(* IEC 61131-3 sources: 2026_Projet_YGO_ExcavatriceDragage/CODE/H_TREUILS_BENNE, 13 files *)

(* ---- FB_BucketCmdArbitration.st ---- *)
(* ═══════════════════════════════════════════════════════════════
   🪣 FB_BucketCmdArbitration — Arbitrage de commande benne
   ───────────────────────────────────────────────────────────────
   🎯 Rôle : Arbitrer la source de commande benne (boutons IHM /
       séquencement couplé both / demande cycle selon le mode) et produire
       les commandes arbitrées (ouverture, fermeture, contacteur Kobold).
   🔌 FB d'arbitrage (non-mouvement) : ne porte ni SafeStop ni StartStop
       de sécurité — il produit la commande logique, la safety reste dans
       FB_Bucket / FB_Safety_Winch.
   📄 Doc : DOC/AF/AF_Partie-10_Fonction_Winch_v2.1.md
   🔒 Bit-identique à l'ancien PRG_04 §1/§2 (refactor POO §5 : décision dans
       le FB, plus dans le PRG). Symétrique à FB_WinchCmdArbitrationM1/M2.
   ═══════════════════════════════════════════════════════════════ *)

FUNCTION_BLOCK FB_BucketCmdArbitration
VAR_INPUT
    Enable    : BOOL;  // --> [CMD] Autorisation FB (TRUE=arbitre actif)
    Auth      : ST_Modes_Autorisations;          // --> [CMD] Autorisations mode (Mode, gating séquencement couplé)
    ReqBucket : ST_ProgramBucketRequest;            // --> [REQ] Demande cycle benne (SEMI_AUTO)
    IHM       : ST_fbBucketCmdArbitration_IHM;      // --> [CMD] Boutons IHM benne (BtnOpen/BtnClose)
    Context   : ST_fbBucketCmdArbitration_Context;   // --> [STAT] Gating séquencement couplé benne
END_VAR
VAR_OUTPUT
    Ready     : BOOL;  // <-- [STAT] FB prêt à arbitrer (Enable)
    CmdOpen_IHM  : BOOL;  // <-- [CMD] Commande ouverture benne arbitrée
    CmdClose_IHM : BOOL;  // <-- [CMD] Commande fermeture benne arbitrée
    KoboldContactorCmdArbitrated : BOOL;  // <-- [CMD] Ordre contacteur capteur fond Kobold arbitré
    WinchBothDiveBucketOpenArmed    : BOOL;  // <-- [STAT] Séquencement couplé : descente benne ouverte armé
    WinchBothAscentBucketCloseArmed : BOOL;  // <-- [STAT] Séquencement couplé : montée benne fermée armé
END_VAR

// === IMPLEMENTATION ===

Ready := Enable;

IF NOT Enable THEN
    CmdOpen_IHM  := FALSE;
    CmdClose_IHM := FALSE;
    KoboldContactorCmdArbitrated := FALSE;
    WinchBothDiveBucketOpenArmed    := FALSE;
    WinchBothAscentBucketCloseArmed := FALSE;
ELSE
    // ── Règle absolue en pilotage both normal (bit-identique PRG_04 §1) ──
    // Descente autorisée UNIQUEMENT benne ouverte, montée UNIQUEMENT benne fermée.
    // T248 : une fois la phase couplée VERROUILLÉE (benne amenée dans l'état requis pour
    // ce maintien joystick), on n'arme plus dive-open / ascent-close -> la perte de
    // l'état ouvert/fermé EN MOUVEMENT ne relance aucune correction benne et ne bloque
    // plus le mouvement couplé ("descente/montée interdite" fantôme).
    WinchBothDiveBucketOpenArmed := Context.TglEnableCoupledBucketSequencing
        AND (Auth.Mode <> E_Mode.SEMI_AUTO)
        AND NOT Context.CoupledPhaseLocked
        AND Context.MotionActive AND Context.ReqDescend
        AND NOT Context.BucketIsOpen;
    WinchBothAscentBucketCloseArmed := Context.TglEnableCoupledBucketSequencing
        AND (Auth.Mode <> E_Mode.SEMI_AUTO)
        AND NOT Context.CoupledPhaseLocked
        AND Context.MotionActive AND Context.ReqAscent
        AND NOT Context.BucketIsClosed;

    // ── Ouverture benne : bouton IHM OU séquencement couplé descente benne ouverte
    //    OU demande cycle (bit-identique PRG_04 §2) ──
    CmdOpen_IHM := IHM.BtnOpen OR WinchBothDiveBucketOpenArmed OR ReqBucket.ReqOpen;

    // ── Fermeture benne : demande cycle > séquencement couplé montée benne fermée
    //    > bouton IHM (bit-identique PRG_04 §1) ──
    IF ReqBucket.ReqClose THEN
        CmdClose_IHM := TRUE;
    ELSIF WinchBothAscentBucketCloseArmed THEN
        CmdClose_IHM := TRUE;
    ELSE
        CmdClose_IHM := IHM.BtnClose;
    END_IF;

    // ── Contacteur Kobold : demande cycle (source unique PRG_03, bit-identique PRG_04 §1) ──
    KoboldContactorCmdArbitrated := ReqBucket.ReqKoboldMeasureEnable;
END_IF;

END_FUNCTION_BLOCK

(* ---- FB_DriftGuard.st ---- *)
(* =======================================================================
   📐 FB_DriftGuard — Détection de dérive de position sous armement
   ───────────────────────────────────────────────────────────────
   🎯 Rôle : Capture position de référence et détection de dérive anormale
   📄 Doc métier : DOC/AF/AF_Partie-10_Fonction_Winch_v2.1.md
   🔌 Interface : Brique interne de sécurité (compose FB_Safety_Winch)
   🔒 Sécurité : Détection de mouvement non commandé et glissement
   ======================================================================= *)

FUNCTION_BLOCK PUBLIC FB_DriftGuard
VAR_INPUT
    // === COMMANDES ET SEUILS ===
    Arm                             : BOOL;                           // --> [CMD] Condition d'armement de la surveillance
    PositionM                       : REAL;                           // --> [HW] Position courante a surveiller (m)
    ToleranceM                      : REAL;                           // --> [CFG] Tolerance de derive maximale autorisee (m)
END_VAR
VAR_OUTPUT
    // === MESURES ET ETATS ===
    RefPosM                         : REAL;                           // <-- [DIAG] Position de reference capturee a l'armement (m)
    DriftM                          : REAL;                           // <-- [DIAG] Derive absolue courante (m)
    Violation                       : BOOL;                           // <-- [STAT] Alarme derive maximale depassee
END_VAR
VAR
    // === VARIABLES LOCALES INTERNES ===
    WasArmed                        : BOOL;                           // . [LOC] Memoire etat armement cycle precedent
END_VAR

// === IMPLEMENTATION (à coller dans le corps ST du POU FB_DriftGuard) ===

IF Arm THEN
    IF NOT WasArmed THEN
        RefPosM := PositionM;   // Capture au 1er cycle armé uniquement
        WasArmed := TRUE;
    END_IF;
    DriftM := ABS(PositionM - RefPosM);
    Violation := DriftM > ToleranceM;
ELSE
    WasArmed := FALSE;
    DriftM := 0.0;
    Violation := FALSE;
END_IF;

(* ---- FB_SpeedStep.st ---- *)
(* =======================================================================
   FB_SpeedStep — Décodeur palier vers contacteurs
   Rôle : applique les bornes de palier puis lit la table contacteurs.
   Le calcul de la consigne discrète est fait par le producteur amont.
   ======================================================================= *)

{attribute 'qualified_only'}
{attribute 'hide_all_locals'}

FUNCTION_BLOCK PUBLIC FB_SpeedStep
VAR_INPUT
    Enable                          : BOOL;
    SpeedStepReq                    : INT := 0;                       // --> [CMD] Palier demandé (0..5)
    Table                           : ST_SpeedStepTable;              // --> [CFG] Table contacteurs propre au treuil
    MinStepNumber                   : INT := 1;                       // --> [CFG] Plancher palier, rétro-compatible
    MaxStepNumber                   : INT := 5;                       // --> [CFG] Plafond palier atteignable
END_VAR
VAR_OUTPUT
    StepNumber                      : INT;                            // <-- [STAT] Palier actif (0..5)
    Contactor1                      : BOOL;                           // <-- [ACT] Ordre contacteur vitesse palier 1
    Contactor2                      : BOOL;                           // <-- [ACT] Ordre contacteur vitesse palier 2
    Contactor3                      : BOOL;                           // <-- [ACT] Ordre contacteur vitesse palier 3
    Contactor4                      : BOOL;                           // <-- [ACT] Ordre contacteur vitesse palier 4
    ConfigError                     : BOOL;                           // <-- [DIAG] Table de paliers invalide
    ConfigErrorId                   : WORD;                           // <-- [DIAG] Bitfield erreur table
END_VAR
VAR
    _ConfigValid                    : BOOL;
    _ConfigErrorIdInt               : WORD;
    _MaxStepClamped                 : INT;
    _MinStepClamped                 : INT;
END_VAR

{region "§0 Bornes et validation table"}
// Le plafond est borné avant le plancher : si le plancher demandé dépasse le
// plafond de sécurité, celui-ci garde la priorité.
_MaxStepClamped := LIMIT(1, MaxStepNumber, 5);
_MinStepClamped := LIMIT(1, MinStepNumber, _MaxStepClamped);

// Les seuils restent validés pour conserver le diagnostic table historique.
// Ils ne participent plus au calcul du palier dans ce FB.
_ConfigValid := TRUE;
_ConfigErrorIdInt := 16#0000;
IF NOT (Table.StepThreshold_Pct[1] < Table.StepThreshold_Pct[2] AND
        Table.StepThreshold_Pct[2] < Table.StepThreshold_Pct[3] AND
        Table.StepThreshold_Pct[3] < Table.StepThreshold_Pct[4] AND
        Table.StepThreshold_Pct[4] < Table.StepThreshold_Pct[5]) THEN
    _ConfigValid := FALSE;
    _ConfigErrorIdInt := _ConfigErrorIdInt OR 16#0001;
END_IF;
IF (Table.StepThreshold_Pct[1] < 0.0) OR (Table.StepThreshold_Pct[5] > 100.0) THEN
    _ConfigValid := FALSE;
    _ConfigErrorIdInt := _ConfigErrorIdInt OR 16#0001;
END_IF;
ConfigErrorId := _ConfigErrorIdInt;
ConfigError := (ConfigErrorId <> 16#0000);
{endregion}

{region "§1 Gate"}
// Relâche ou table invalide : aucun plancher ne peut maintenir un contacteur.
IF (NOT Enable) OR (NOT _ConfigValid) OR (SpeedStepReq <= 0) THEN
    StepNumber := 0;
    Contactor1 := FALSE; Contactor2 := FALSE; Contactor3 := FALSE; Contactor4 := FALSE;
    RETURN;
END_IF;
{endregion}

{region "§2 Clamp et table contacteurs"}
// Le plancher agit sur la cible. StepNumber ne reçoit jamais directement
// MinStepNumber ; LIMIT final garantit la plage 1..5 après le plafond.
StepNumber := LIMIT(_MinStepClamped, SpeedStepReq, _MaxStepClamped);

CASE StepNumber OF
    1:  Contactor1 := Table.P1R1; Contactor2 := Table.P1R2; Contactor3 := Table.P1R3; Contactor4 := Table.P1R4;
    2:  Contactor1 := Table.P2R1; Contactor2 := Table.P2R2; Contactor3 := Table.P2R3; Contactor4 := Table.P2R4;
    3:  Contactor1 := Table.P3R1; Contactor2 := Table.P3R2; Contactor3 := Table.P3R3; Contactor4 := Table.P3R4;
    4:  Contactor1 := Table.P4R1; Contactor2 := Table.P4R2; Contactor3 := Table.P4R3; Contactor4 := Table.P4R4;
    5:  Contactor1 := Table.P5R1; Contactor2 := Table.P5R2; Contactor3 := Table.P5R3; Contactor4 := Table.P5R4;
ELSE
    // Défense en profondeur face à une divergence type/outil.
    StepNumber := 0;
    Contactor1 := FALSE; Contactor2 := FALSE; Contactor3 := FALSE; Contactor4 := FALSE;
END_CASE;
{endregion}

END_FUNCTION_BLOCK

(* ---- FB_SyncContactor.st ---- *)
(* =======================================================================
   🔀 FB_SyncContactor — Coherence commandes/contacteurs M1/M2
   ───────────────────────────────────────────────────────────────
   🎯 Rôle : Detecter une discordance entre les commandes/contacteurs des
      2 treuils (sens + paliers). Independante des codeurs — surveillable
      meme si les codeurs sont bypasses.
   🔌 Interface : Bloc de surveillance transverse (1..N instances : requetes
      amont dans FB_WinchSync, sorties physiques finales dans PRG_06).
   🔒 Polarite : ContactorMismatch = TRUE si discordance confirmee (debounce).
      Reponse GRADUEE : ContactorMismatch (niveau 1, filtre MismatchDebounce)
      -> SafeStop ; ContactorMismatchEscalated (niveau 2, si la discordance
      tient CST_SyncEscalationTime) -> escalade PowerCutOff.
   ⚖️ Concordance ACTIVE des que les 2 treuils sont commandes (relais ou
      contacteur) OU en mode synchronisme (SyncEnable). Seul BypassGlobal
      neutralise.
   📄 Doc : DOC/AF/AF_Partie-10_Fonction_Winch_v2.1.md
   ======================================================================= *)

FUNCTION_BLOCK PUBLIC FB_SyncContactor
VAR_INPUT
    // === COMMANDES ET CONSIGNES ===
    Enable                          : BOOL;                           // --> [CMD] Validation surveillance globale
    Reset                           : BOOL;                           // --> [CMD] Acquittement defaut sur front
    SyncEnable                      : BOOL;                           // --> [CMD] Autorisation utilisateur synchro

    // === COMMANDES ET FEEDBACKS ACTIONS ===
    RelayFwdM1                      : BOOL;                           // --> [HW] Feedback/Ordre montee M1
    RelayFwdM2                      : BOOL;                           // --> [HW] Feedback/Ordre montee M2
    RelayRevM1                      : BOOL;                           // --> [HW] Feedback/Ordre descente M1
    RelayRevM2                      : BOOL;                           // --> [HW] Feedback/Ordre descente M2
    Contactor1_M1                   : BOOL;                           // --> [HW] Contacteur palier 1 M1
    Contactor1_M2                   : BOOL;                           // --> [HW] Contacteur palier 1 M2
    Contactor2_M1                   : BOOL;                           // --> [HW] Contacteur palier 2 M1
    Contactor2_M2                   : BOOL;                           // --> [HW] Contacteur palier 2 M2
    Contactor3_M1                   : BOOL;                           // --> [HW] Contacteur palier 3 M1
    Contactor3_M2                   : BOOL;                           // --> [HW] Contacteur palier 3 M2
    Contactor4_M1                   : BOOL;                           // --> [HW] Contacteur palier 4 M1
    Contactor4_M2                   : BOOL;                           // --> [HW] Contacteur palier 4 M2

    // === BYPASSES ET SIMULATION ===
    BypassGlobal                    : BOOL := FALSE;                  // --> [TST] Neutralise la surveillance contacteurs
    DescentStep45Permit             : BOOL := FALSE;                  // --> [CMD] Autorise uniquement le profil descente M1=P4 / M2=P5
    SpeedStepTable                  : ST_SpeedStepTable;              // --> [CFG] Table officielle paliers -> contacteurs
END_VAR
VAR_OUTPUT
    // === RESULTAT (reponse graduee) ===
    ContactorMismatch               : BOOL;                           // <-- [SAFE] Niveau 1 : discordance commande/contacteurs confirmee (debounce) -> SafeStop
    ContactorMismatchEscalated      : BOOL;                           // <-- [SAFE] Niveau 2 : discordance persistante -> escalade PowerCutOff
    CommandsCoherent                : BOOL;                           // <-- [STAT] TRUE si le vecteur instantane est coherent ou derogation T291-A exacte
    DescentStep45Matched            : BOOL;                           // <-- [STAT] TRUE si le profil M1=P4 / M2=P5 est exactement reconnu
    Diag                            : ST_SyncContactorDiag;           // <-- [DIAG] Detail : quel contacteur diverge + niveau atteint
END_VAR
VAR CONSTANT
    MismatchDebounce                : TIME := T#500ms;                // Filtre transitoires/rampes avant de confirmer la discordance (niveau 1)
    CST_SyncEscalationTime          : TIME := T#3s;                   // Discordance confirmee tenue au-dela de ce delai -> escalade (niveau 2)
END_VAR
VAR
    // === DETECTEURS ET TIMERS INTERNES ===
    MismatchTimer                   : TON;                            // . [LOC] Tempo filtrage incoherence (niveau 1)
    EscalationTimer                 : TON;                            // . [LOC] Tempo escalade (niveau 2)

    // === VARIABLES LOCALES INTERNES ===
    MismatchActive                  : BOOL;                           // . [LOC] Discordance instantanee (avant debounce)
    BothCommanded                   : BOOL;                           // . [LOC] Les 2 treuils sont commandes (relais ou contacteur)
    DescentStep4M1                  : BOOL;                           // . [LOC] M1 en descente avec vecteur table P4 exact
    DescentStep5M2                  : BOOL;                           // . [LOC] M2 en descente avec vecteur table P5 exact
END_VAR

{region "§1 Gate neutralisation"}
// 🛑 1. GATE
IF NOT Enable OR BypassGlobal THEN
    ContactorMismatch := FALSE;
    ContactorMismatchEscalated := FALSE;
    CommandsCoherent := FALSE;
    DescentStep45Matched := FALSE;
    MismatchActive := FALSE;
    BothCommanded := FALSE;
    DescentStep4M1 := FALSE;
    DescentStep5M2 := FALSE;
    MismatchTimer(IN := FALSE);
    EscalationTimer(IN := FALSE);
    Diag.RelayFwdMismatch := FALSE;
    Diag.RelayRevMismatch := FALSE;
    Diag.Step1Mismatch := FALSE;
    Diag.Step2Mismatch := FALSE;
    Diag.Step3Mismatch := FALSE;
    Diag.Step4Mismatch := FALSE;
    Diag.MismatchLevel := 0;
    RETURN;
END_IF;
{endregion}

{region "§2 Detection discordance + diagnostic decode"}
// 🔍 2. COHÉRENCE DES COMMANDES SÉCURITÉ — verifie que les commandes envoyees
// aux deux treuils sont identiques (sens et contacteurs).
// Concordance ACTIVE des que les 2 treuils sont commandes (relais ou contacteur)
// OU en mode synchronisme (SyncEnable).
BothCommanded := (RelayFwdM1 OR RelayRevM1 OR Contactor1_M1 OR Contactor2_M1
                  OR Contactor3_M1 OR Contactor4_M1)
             AND (RelayFwdM2 OR RelayRevM2 OR Contactor1_M2 OR Contactor2_M2
                  OR Contactor3_M2 OR Contactor4_M2);

// Diagnostic decode : quel(s) contacteur(s) diverge(nt) (bits nommes, plusieurs possibles).
Diag.RelayFwdMismatch := (BothCommanded OR SyncEnable) AND (RelayFwdM1 <> RelayFwdM2);
Diag.RelayRevMismatch := (BothCommanded OR SyncEnable) AND (RelayRevM1 <> RelayRevM2);
Diag.Step1Mismatch    := (BothCommanded OR SyncEnable) AND (Contactor1_M1 <> Contactor1_M2);
Diag.Step2Mismatch    := (BothCommanded OR SyncEnable) AND (Contactor2_M1 <> Contactor2_M2);
Diag.Step3Mismatch    := (BothCommanded OR SyncEnable) AND (Contactor3_M1 <> Contactor3_M2);
Diag.Step4Mismatch    := (BothCommanded OR SyncEnable) AND (Contactor4_M1 <> Contactor4_M2);

DescentStep4M1 := RelayRevM1 AND NOT RelayFwdM1
                  AND (Contactor1_M1 = SpeedStepTable.P4R1)
                  AND (Contactor2_M1 = SpeedStepTable.P4R2)
                  AND (Contactor3_M1 = SpeedStepTable.P4R3)
                  AND (Contactor4_M1 = SpeedStepTable.P4R4);
DescentStep5M2 := RelayRevM2 AND NOT RelayFwdM2
                  AND (Contactor1_M2 = SpeedStepTable.P5R1)
                  AND (Contactor2_M2 = SpeedStepTable.P5R2)
                  AND (Contactor3_M2 = SpeedStepTable.P5R3)
                  AND (Contactor4_M2 = SpeedStepTable.P5R4);
DescentStep45Matched := DescentStep45Permit
                        AND NOT RelayFwdM2
                        AND NOT RelayFwdM1
                        AND DescentStep4M1
                        AND DescentStep5M2;

IF DescentStep45Matched THEN
    Diag.Step1Mismatch := FALSE;
    Diag.Step2Mismatch := FALSE;
    Diag.Step3Mismatch := FALSE;
    Diag.Step4Mismatch := FALSE;
END_IF;

MismatchActive := Diag.RelayFwdMismatch OR Diag.RelayRevMismatch
    OR Diag.Step1Mismatch OR Diag.Step2Mismatch
    OR Diag.Step3Mismatch OR Diag.Step4Mismatch;
CommandsCoherent := NOT MismatchActive;

// Niveau 1 : discordance confirmee apres MismatchDebounce.
MismatchTimer(IN := MismatchActive, PT := MismatchDebounce);
ContactorMismatch := MismatchTimer.Q;

// Niveau 2 : la discordance confirmee tient au-dela de CST_SyncEscalationTime.
EscalationTimer(IN := ContactorMismatch, PT := CST_SyncEscalationTime);
ContactorMismatchEscalated := EscalationTimer.Q;

// Niveau publie.
IF ContactorMismatchEscalated THEN
    Diag.MismatchLevel := 2;
ELSIF ContactorMismatch THEN
    Diag.MismatchLevel := 1;
ELSE
    Diag.MismatchLevel := 0;
END_IF;
{endregion}

END_FUNCTION_BLOCK

(* ---- FB_Winch.st ---- *)
(* =======================================================================
   🪝 FB_Winch — Directeur d'un treuil individuel (M1 / M2)
   ───────────────────────────────────────────────────────────────
   🎯 Rôle : Pilotage d'un treuil individuel (contacteurs de sens et de vitesse)
   📄 Doc métier : DOC/AF/AF_Partie-10_Fonction_Winch_v2.1.md
   🔌 Interface : FB de mouvement (Enable, SafeStop, RunRequest via WinchRequest)
   🔒 Sécurité : Interlock inversion de sens et gestion des autorisations
   🔧 Interface plate → structs (WinchRequest / Sensors / Config),
      logique interne conservée (comportement bit-identique).
   ======================================================================= *)

FUNCTION_BLOCK PUBLIC FB_Winch
VAR_INPUT
    // === COMMANDES ET CONSIGNES ===
    Enable                          : BOOL;                           // --> [CMD] Autorisation generale FB (TRUE=Autorise)
    Reset                           : BOOL;                           // --> [CMD] Acquittement defaut (front)
    PowerContactorEngaged           : BOOL;                           // --> [SAFE] Statut contacteur de ligne / puissance

    // === REQUÊTE D'AXE (struct) ===
    WinchRequest                    : ST_fbWinch_Req;                  // --> [REQ] RunRequest + 2 bits de sens, palier et limites

    // === MESURES ET FEEDBACKS (struct) ===
    Sensors                         : ST_fbWinch_Sensors;             // --> [HW] Position, referencement, contacteurs, vitesse

    // === CONFIGURATION STATIQUE (struct) ===
    Config                          : ST_fbWinch_Cfg;                 // --> [CFG] Table paliers, delais, ralentissement

    // === SECOURS ET PERMIS DE SÉCURITÉ ===
    SafeStop                        : BOOL;                           // --> [SAFE] Arret rapide de securite
    DescendPermit                   : BOOL := FALSE;                 // --> [SAFE] Permis de descente (mou de cable)
    AscentPermit                    : BOOL := FALSE;                 // --> [SAFE] Permis de montee (fin de course haut)

    // === BYPASSES ET SIMULATION ===
    BypassContactorCheck            : BOOL;                           // --> [TST] Bypass diagnostic contacteurs (simu)
    BypassGlobal                    : BOOL;                           // --> [TST] Force ErrorId=0, ignore erreurs
END_VAR
VAR_OUTPUT
    // === ETATS IEC ET SYNOPTIQUE ===
    Ready                           : BOOL;                           // <-- [STAT] FB pret a fonctionner
    // 🧩 Statut transverse (forme cible ST_Fault)
    Fault                           : ST_Fault;

    // === ORDRES ACTIONNEURS (CONTACTEURS) ===
    RelayFwd                        : BOOL;                           // <-- [ACT] Ordre contacteur sens montee
    RelayRev                        : BOOL;                           // <-- [ACT] Ordre contacteur sens descente
    Contactor1                      : BOOL;                           // <-- [ACT] Ordre contacteur vitesse palier 1
    Contactor2                      : BOOL;                           // <-- [ACT] Ordre contacteur vitesse palier 2
    Contactor3                      : BOOL;                           // <-- [ACT] Ordre contacteur vitesse palier 3
    Contactor4                      : BOOL;                           // <-- [ACT] Ordre contacteur vitesse palier 4

    // === DIAGNOSTICS ET MESURES ===
    RequestedStep                   : INT;                            // <-- [DIAG] Palier brut calcule par SpeedStep
    StepNumber                      : INT;                            // <-- [DIAG] Palier metier temporise actif
    BusinessStepDelayElapsed        : TIME;                           // <-- [DIAG] Ecoule tempo metier palier
    SpeedGuardLimited               : BOOL;                           // <-- [DIAG] Statut limitation par garde-fou
    ContactorsCheck                 : ST_ContactorCheck;              // <-- [DIAG] Diagnostic concorde contacteurs
    InTopSlowdownZone               : BOOL;                           // <-- [DIAG] Zone de ralentissement haut active
    InBottomSlowdownZone            : BOOL;                           // <-- [DIAG] Zone de ralentissement bas active
    CommandedAscent                 : BOOL;                           // <-- [DIAG] Sens interne mémorisé : montée
    CommandedDescend                : BOOL;                           // <-- [DIAG] Sens interne mémorisé : descente
    RequestConflict                 : BOOL;                           // <-- [DIAG] Double demande de sens détectée
    DirectionChangeDelayElapsed     : TIME;                           // <-- [DIAG] Ecoule delai changement de sens
    DirectionChangePending          : BOOL;                           // <-- [DIAG] Changement de sens en attente

    // === INTENTION DE MAINTIEN DU CONTACTEUR DE SENS (§3bis) ===
    SenseHoldRequest                : BOOL;                           // <-- [ACT] Demande a la barriere finale de TENIR le contacteur de sens apres chute de palier a 0 (inertie moteur), bornee par T_hold_internal
END_VAR
VAR
    // === SOUS-INSTANCES FB ===
    SpeedStep                       : FB_SpeedStep;                   // * [INST] Decodage paliers vitesse
    DirectionInterlock              : FB_WinchDirectionInterlock;     // * [INST] Interlock changement de sens (D18)
    StepShaper                      : FB_WinchStepShaper;             // * [INST] Cadencement de palier (D10)

    // === DETECTEURS ET TIMERS INTERNES ===
    ResetEdge                       : R_TRIG;                         // . [LOC] Detecteur front montant Reset
    EnableRisingEdge                : R_TRIG;                         // . [LOC] Detecteur front montant Enable (D18)
    TonContactorsDropped            : TON;                            // . [LOC] Temporisation retombee contacteurs

    // === VARIABLES LOCALES CALCULÉES ===
    AllContactorsCommandedOff       : BOOL;                           // . [LOC] Tous contacteurs commandes a FALSE
    RampTargetStep                  : INT;                            // . [LOC] Palier demandé par l'arbitrage amont
    EffectiveSafeStop               : BOOL;                           // . [LOC] SafeStop effectif incluant permis
    DirectionConflict               : BOOL;                           // . [LOC] Les deux demandes de sens sont actives
    ActiveMaxStep                   : INT;                            // . [LOC] Plafond palier actif dynamique
    EffectiveStepRampDelay          : TIME;                           // . [LOC] Cadence palier selon sens, distincte interlock

    // === MAINTIEN DU CONTACTEUR DE SENS (§3bis) ===
    SenseHoldTimer                  : TON;                            // . [LOC] Garde interne T_hold_internal (< MaxSenseHoldTime barriere)
    SenseHoldActiveInt              : BOOL;                           // . [LOC] Maintien de sens interne en cours
    PrevStepNumber                  : INT;                            // . [LOC] Palier temporise du scan precedent (detection chute a 0)
    SenseHoldHardCut                : BOOL;                           // . [LOC] Coupure dure active (interdit tout maintien)

    // Latches défauts
    SpeedStepConfigFaultLatched     : BOOL;

    // Socle défaut
    instFault                       : FB_FaultCore;                   // * [INST] Socle défaut transverse
    instCauses                      : ARRAY[0..15] OF ST_FaultCause;  // . [LOC] Table des causes nommées
END_VAR

// === IMPLEMENTATION ===

{region "§1 Causes & Socle Défaut (évalué en continu)"}
// 🔑 1. FRONTS & REARMEMENT
ResetEdge(CLK := Reset);
EnableRisingEdge(CLK := Enable);

IF ResetEdge.Q OR BypassGlobal THEN
    SpeedStepConfigFaultLatched := FALSE;
    ContactorsCheck.StuckClosed := FALSE;
END_IF;

IF Enable AND SpeedStep.ConfigError THEN
    SpeedStepConfigFaultLatched := TRUE;
END_IF;

// FB_Safety_Winch est l'unique proprietaire de la detection contacteur colle.
// FB_Winch conserve le champ public pour compatibilite IHM/Troubleshooting,
// mais ne produit plus ce defaut.
instCauses[1].Active   := FALSE;
instCauses[1].Latching := TRUE;
instCauses[1].Texte    := 'Contacteur colle gere par FB_Safety_Winch ';

instCauses[2].Active   := SpeedStepConfigFaultLatched;
instCauses[2].Latching := TRUE;
instCauses[2].Texte    := 'Configuration table des paliers vitesse invalide';

// Appel du socle de défaut
instFault(Enable := Enable, Reset := Reset, Causes := instCauses);
Fault := instFault.Fault;
{endregion}

{region "§2 Gate neutralisation"}
// 🛑 2. GATE
IF NOT Enable THEN
    SpeedStep(Enable := FALSE, SpeedStepReq := 0, Table := Config.SpeedStepTable);
    DirectionInterlock(Enable := FALSE, EnableRising := FALSE, Reset := Reset, ReqAscent := FALSE, ReqDescend := FALSE,
                       ChangeDelayAscent := Config.DirectionInterlockDelayAscent,
                       ChangeDelayDescent := Config.DirectionInterlockDelayDescent);
    StepShaper(Enable := FALSE, TargetStep := 0, StepRampDelay := Config.StepRampDelayAscent);
    RelayFwd := FALSE;
    RelayRev := FALSE;
    Contactor1 := FALSE; Contactor2 := FALSE; Contactor3 := FALSE; Contactor4 := FALSE;
    RequestedStep := 0;
    StepNumber := StepShaper.ShapedStep;
    CommandedAscent := DirectionInterlock.CommandedAscent;
    CommandedDescend := DirectionInterlock.CommandedDescend;
    RequestConflict := DirectionInterlock.RequestConflict;
    DirectionChangePending := DirectionInterlock.DirectionChangePending;
    TonContactorsDropped(IN := FALSE);
    ContactorsCheck.Command := FALSE;
    ContactorsCheck.Feedback := NOT Sensors.ContactorsAllOff;
    InTopSlowdownZone := FALSE;
    InBottomSlowdownZone := FALSE;
    // §3bis : coupure dure -> aucun maintien de sens possible, etat interne purge.
    SenseHoldRequest := FALSE;
    SenseHoldActiveInt := FALSE;
    SenseHoldTimer(IN := FALSE, PT := T#900ms);
    PrevStepNumber := 0;
    Ready := FALSE;
    RETURN;
END_IF;

Ready := Enable AND NOT Fault.Latched;
{endregion}

{region "§3 Permis et zones de ralentissement"}
DirectionConflict := WinchRequest.ReqAscent AND WinchRequest.ReqDescend;
EffectiveSafeStop := SafeStop OR DirectionConflict
                     OR (WinchRequest.ReqAscent AND NOT AscentPermit)
                     OR (WinchRequest.ReqDescend AND NOT DescendPermit);

InTopSlowdownZone := Sensors.Homed AND NOT Sensors.HomingSuspect AND (Sensors.CablePosM >= (WinchRequest.TopLimitM - Config.SlowdownDistanceTop_M));
InBottomSlowdownZone := Sensors.Homed AND NOT Sensors.HomingSuspect AND (Sensors.CablePosM <= (WinchRequest.BottomLimitM + Config.SlowdownDistanceBottom_M));

IF WinchRequest.ReqAscent AND NOT WinchRequest.ReqDescend THEN
    ActiveMaxStep := WinchRequest.MaxStepUp;
    IF InTopSlowdownZone THEN
        ActiveMaxStep := MIN(ActiveMaxStep, Config.SlowdownMaxStep);
    END_IF;
ELSIF WinchRequest.ReqDescend AND NOT WinchRequest.ReqAscent THEN
    ActiveMaxStep := WinchRequest.MaxStepDown;
    IF InBottomSlowdownZone THEN
        ActiveMaxStep := MIN(ActiveMaxStep, Config.SlowdownMaxStep);
    END_IF;
ELSE
    ActiveMaxStep := WinchRequest.MaxStepUp;
END_IF;

IF WinchRequest.HomingApproachActive THEN
    ActiveMaxStep := 1;
END_IF;
{endregion}

{region "§4 Interlock direction"}
// 🔀 4. INTERLOCK DIRECTION (extrait dans FB_WinchDirectionInterlock, D18)
DirectionInterlock(
    Enable := (StepNumber = 0) AND Sensors.ContactorsAllOff,
    EnableRising := EnableRisingEdge.Q,
    Reset := Reset,
    ReqAscent := WinchRequest.ReqAscent,
    ReqDescend := WinchRequest.ReqDescend,
    ChangeDelayAscent := Config.DirectionInterlockDelayAscent,
    ChangeDelayDescent := Config.DirectionInterlockDelayDescent
);
CommandedAscent := DirectionInterlock.CommandedAscent;
CommandedDescend := DirectionInterlock.CommandedDescend;
RequestConflict := DirectionInterlock.RequestConflict;
DirectionChangePending := DirectionInterlock.DirectionChangePending;
DirectionChangeDelayElapsed := DirectionInterlock.DelayElapsed;
{endregion}

{region "§5 Paliers vitesse et contacteurs"}
// -B : la consigne est désormais un PALIER discret (WinchRequest.SpeedStepReq,
// 1..5, 0 = arrêt) produit par l'arbitrage. Plus de décodage %→palier ici.
IF DirectionChangePending OR NOT (WinchRequest.ReqAscent OR WinchRequest.ReqDescend) OR EffectiveSafeStop OR NOT WinchRequest.RunRequest THEN
    RampTargetStep := 0;
ELSE
    RampTargetStep := WinchRequest.SpeedStepReq;
END_IF;

SpeedStep(
    Enable := (RampTargetStep > 0),
    SpeedStepReq := RampTargetStep,
    Table := Config.SpeedStepTable,
    MaxStepNumber := ActiveMaxStep
);
RequestedStep := SpeedStep.StepNumber;

// 🛡️ Garde-fou vitesse : bride le palier demande si la vitesse n'est pas stable
// (SpeedGuardReady=FALSE -> palier 1) ou si la bande mesuree est inferieure au
// palier demande (pas de passage aux paliers superieurs sans vitesse confirmee).
SpeedGuardLimited := FALSE;
IF Sensors.SpeedGuardEnable THEN
    IF NOT Sensors.SpeedGuardReady THEN
        IF RequestedStep > 1 THEN
            RequestedStep := 1;
            SpeedGuardLimited := TRUE;
        END_IF;
    ELSIF (Sensors.MeasuredSpeedBand >= 1) AND (Sensors.MeasuredSpeedBand <= 5) AND (RequestedStep > Sensors.MeasuredSpeedBand) THEN
        RequestedStep := Sensors.MeasuredSpeedBand;
        SpeedGuardLimited := TRUE;
    END_IF;
END_IF;

// 🤿 Plancher palier descente -- plongee Kobold.
// Injecte MinStepDown sur la CIBLE (RequestedStep, consommee par le shaper ci-dessous),
// JAMAIS sur StepNumber directement. Actif uniquement en descente commandee
// ET NON bloquee par un arret/permis (NOT EffectiveSafeStop) : un permis descente FALSE
// doit interdire physiquement le mouvement, sans re-atterrissage du plancher.
// Le sens doit aussi etre deja adopte : pendant DirectionChangePending, le
// StepNumber doit rester a 0 afin que le temps mort d'inversion puisse s'ecouler.
// (RunRequest AND ReqDescend) : relache joystick (RunRequest=FALSE) -> aucun plancher,
// l'arret franc RequestedStep=0 / RampTargetStep=0 est preserve.
// Regle d'agregation : le PLAFOND GAGNE -- si le plancher depasse le plafond courant
// ActiveMaxStep (ex. SlowdownMaxStep -> palier 1 en bordure basse), on borne au plafond.
IF WinchRequest.RunRequest AND WinchRequest.ReqDescend AND NOT WinchRequest.ReqAscent
   AND (WinchRequest.MinStepDown > 0) AND NOT EffectiveSafeStop
   AND NOT DirectionChangePending AND CommandedDescend THEN
    IF RequestedStep < WinchRequest.MinStepDown THEN
        RequestedStep := WinchRequest.MinStepDown;
    END_IF;
    IF RequestedStep > ActiveMaxStep THEN
        RequestedStep := ActiveMaxStep;
    END_IF;
END_IF;

// ⚙️ Cadencement de palier (extrait dans FB_WinchStepShaper, D10).
// Les deux cadences historiques sont preservees sans reutiliser les delais
// d'interlock direction : 1 s en montee, 500 ms en descente.
IF CommandedDescend THEN
    EffectiveStepRampDelay := Config.StepRampDelayDescent;
ELSE
    EffectiveStepRampDelay := Config.StepRampDelayAscent;
END_IF;
StepShaper(
    Enable := Enable,
    TargetStep := RequestedStep,
    StepRampDelay := EffectiveStepRampDelay
);
StepNumber := StepShaper.ShapedStep;
BusinessStepDelayElapsed := StepShaper.StepDelayElapsed;

IF StepNumber > 0 AND CommandedAscent THEN
    RelayFwd := TRUE;
    RelayRev := FALSE;
ELSIF StepNumber > 0 AND CommandedDescend THEN
    RelayFwd := FALSE;
    RelayRev := TRUE;
ELSE
    RelayFwd := FALSE;
    RelayRev := FALSE;
END_IF;

// 🛡️ FIX contacteurs (audit CONTACTEURS_2026-08-31) + SOLUTION : ré-émettre les
// contacteurs depuis FB_SpeedStep (décodage TABLE ST_SpeedStepTable cumulatif :
// P1=0, P2={K1}, P3={K1,K2}, P4={K1,K2,K3}, P5={K1,K2,K3,K4}) sur le palier SHAPÉ,
// au lieu de l'ancien décodage one-hot exclusif (ContactorN := StepNumber=N) qui
// éteignait les paliers inférieurs et ne couvrait pas le palier 5.
SpeedStep(
    Enable          := (StepNumber > 0),
    SpeedStepReq    := StepNumber,
    Table           := Config.SpeedStepTable,
    MaxStepNumber   := ActiveMaxStep
);
Contactor1 := SpeedStep.Contactor1;
Contactor2 := SpeedStep.Contactor2;
Contactor3 := SpeedStep.Contactor3;
Contactor4 := SpeedStep.Contactor4;

AllContactorsCommandedOff := (NOT RelayFwd) AND (NOT RelayRev)
                             AND (NOT Contactor1) AND (NOT Contactor2) AND (NOT Contactor3) AND (NOT Contactor4);

ContactorsCheck.Command  := NOT AllContactorsCommandedOff;
ContactorsCheck.Feedback := NOT Sensors.ContactorsAllOff;
TonContactorsDropped(IN := FALSE, PT := Config.ContactorFeedbackTimeout);
ContactorsCheck.StuckClosed := FALSE; // force a FALSE (Phase 0) : detection contacteur colle produite par FB_Safety_Winch, re-alimentee a la phase suivante
ContactorsCheck.StuckOpen := FALSE;

IF Fault.Error THEN
    RelayFwd := FALSE;
    RelayRev := FALSE;
    Contactor1 := FALSE; Contactor2 := FALSE; Contactor3 := FALSE; Contactor4 := FALSE;
END_IF;
{endregion}

{region "§5bis Intention de maintien du contacteur de sens (§3bis)"}
// Quand le palier temporise StepNumber vient de retomber a 0 alors qu'un sens etait
// commande, FB_Winch DEMANDE a la barriere finale (FB_WinchOutputInterlock) de TENIR
// le contacteur de sens le temps que le moteur ralentisse (inertie). Borne par
// T_hold_internal (garde interne, < MaxSenseHoldTime de la barriere = T#1s).
// Coupures dures -> retombee immediate, jamais de maintien (SafeStop / defaut / perte
// puissance / NOT Enable geree a la gate §2).
SenseHoldHardCut := (NOT PowerContactorEngaged) OR EffectiveSafeStop OR Fault.Error;

IF SenseHoldHardCut THEN
    SenseHoldActiveInt := FALSE;
ELSIF (PrevStepNumber > 0) AND (StepNumber = 0) AND (CommandedAscent OR CommandedDescend) THEN
    SenseHoldActiveInt := TRUE;   // front de chute de palier a 0 avec sens encore actif
END_IF;

// Maintien interne aligné sur MaxSenseHoldTime de FB_WinchOutputInterlock (T#400ms).
SenseHoldTimer(IN := SenseHoldActiveInt, PT := T#400ms);
IF SenseHoldTimer.Q OR (StepNumber > 0) THEN
    SenseHoldActiveInt := FALSE;  // borne de temps atteinte, ou nouveau mouvement demande
END_IF;

SenseHoldRequest := SenseHoldActiveInt AND NOT SenseHoldHardCut;
PrevStepNumber := StepNumber;
{endregion}

END_FUNCTION_BLOCK

(* ---- FB_Winch_Symmetry.st ---- *)
(* =======================================================================
   ⚖️ FB_Winch_Symmetry — Mesure passive M1/M2
   ───────────────────────────────────────────────────────────────
   🎯 Rôle : Observateur de symétrie et de synchronisme des treuils M1/M2
   📄 Doc métier : DOC/AF/AF_Partie-10_Fonction_Winch_v2.1.md
   🔒 Observateur pur : Aucune ecriture de commande, securite ou mouvement
   ======================================================================= *)

FUNCTION_BLOCK FB_Winch_Symmetry
VAR_INPUT
    // === COMMANDES ET CONSIGNES ===
    Reset                           : BOOL;                           // --> [CMD] Reinitialisation des mesures sur front
    M1CommandActive                 : BOOL;                           // --> [CMD] Commande active sur treuil M1
    M2CommandActive                 : BOOL;                           // --> [CMD] Commande active sur treuil M2
    M1Direction                     : INT;                            // --> [CMD] Sens commande M1 (-1/0/+1)
    M2Direction                     : INT;                            // --> [CMD] Sens commande M2 (-1/0/+1)

    // === FEEDBACKS HARWARE ET FREINS ===
    M1BrakeCmd                      : BOOL;                           // --> [HW] Ordre ouverture frein M1
    M2BrakeCmd                      : BOOL;                           // --> [HW] Ordre ouverture frein M2
    M1BrakeApplied                  : BOOL;                           // --> [HW] Etat frein M1 serre
    M2BrakeApplied                  : BOOL;                           // --> [HW] Etat frein M2 serre

    // === MESURES POSITIONS ET VITESSES ===
    M1Position_M                    : REAL;                           // --> [HW] Position mesuree M1 (m)
    M2Position_M                    : REAL;                           // --> [HW] Position mesuree M2 (m)
    M1Speed_Mps                     : REAL;                           // --> [HW] Vitesse mesuree M1 (m/s)
    M2Speed_Mps                     : REAL;                           // --> [HW] Vitesse mesuree M2 (m/s)
    SyncDeviation_M                 : REAL;                           // --> [HW] Ecart instantane synchro (m)

    // === CONFIGURATION ===
    Config                          : ST_fbWinch_Symmetry_Cfg;           // --> [CFG] Configuration des seuils de symetrie
END_VAR
VAR_OUTPUT
    // === ETATS IEC ET SYNOPTIQUE ===
    SymmetryOk                      : BOOL;                           // <-- [STAT] Symetrie globale conforme aux criteres
    SymmetryValid                   : BOOL;                           // <-- [STAT] Mesure de symetrie valide et calculee
END_VAR
VAR_IN_OUT
    // === STRUCTURES DE DONNÉES PARTAGÉES ===
    Data                            : ST_fbWinch_Symmetry_Data;          // <-> [BUS] Donnees de mesures de symetrie
END_VAR
VAR
    // === SOUS-INSTANCES FB ===
    ResetEdge                       : R_TRIG;                         // * [INST] Detecteur front reinitialisation
    CycleTime                       : FB_CycleTime;                   // * [INST] Calcul du temps de cycle

    // === TIMERS INTERNES ===
    CommandTon                      : TON;                            // . [LOC] Tempo qualification commande stable
    MotionTimer                     : TON;                            // . [LOC] Chronometre de mouvement
    StopTimer                       : TON;                            // . [LOC] Chronometre d'arret

    // === VARIABLES LOCALES CALCULÉES ===
    Comparable                      : BOOL;                           // . [LOC] Conditions de comparaison remplies
    Qualified                       : BOOL;                           // . [LOC] Phase de mesure qualifiee
    PreviousQualified               : BOOL;                           // . [LOC] Etat qualifie cycle precedent
    Stopping                        : BOOL;                           // . [LOC] Phase d'arret en cours
    StartCapturedM1                 : BOOL;                           // . [LOC] Top depart capture M1
    StartCapturedM2                 : BOOL;                           // . [LOC] Top depart capture M2
    StopCapturedM1                  : BOOL;                           // . [LOC] Top arret capture M1
    StopCapturedM2                  : BOOL;                           // . [LOC] Top arret capture M2
    StartMsM1                       : UDINT;                          // . [LOC] Horodatage d'ouverture M1 (ms)
    StartMsM2                       : UDINT;                          // . [LOC] Horodatage d'ouverture M2 (ms)
    ReleaseMsM1                     : UDINT;                          // . [LOC] Temps de desserrage frein M1 (ms)
    ReleaseMsM2                     : UDINT;                          // . [LOC] Temps de desserrage frein M2 (ms)
    ApplyMsM1                       : UDINT;                          // . [LOC] Temps de serrage frein M1 (ms)
    ApplyMsM2                       : UDINT;                          // . [LOC] Temps de serrage frein M2 (ms)
    StopMsM1                        : UDINT;                          // . [LOC] Horodatage d'arret M1 (ms)
    StopMsM2                        : UDINT;                          // . [LOC] Horodatage d'arret M2 (ms)
    StopStartM1_M                   : REAL;                           // . [LOC] Position debut d'arret M1 (m)
    StopStartM2_M                   : REAL;                           // . [LOC] Position debut d'arret M2 (m)
END_VAR

{region "§1 Reset et qualification"}
CycleTime(DefaultValueS := 0.010); ResetEdge(CLK := Reset);
IF ResetEdge.Q THEN Data.DeltaStartDelay_Ms:=0; Data.DeltaBrakeReleaseTime_Ms:=0; Data.DeltaBrakeApplyTime_Ms:=0; Data.DeltaStopDistance_Mm:=0; Data.DeltaStopTime_Ms:=0; Data.MaxSyncDeviation_M:=0.0; END_IF;
Comparable := M1CommandActive AND M2CommandActive AND (M1Direction = M2Direction) AND (M1Direction <> 0);
CommandTon(IN := Comparable, PT := UDINT_TO_TIME(Config.MinimumCommandTime_Ms));
Qualified := CommandTon.Q AND (M1Speed_Mps >= Config.MinimumSpeed_Mps) AND (M2Speed_Mps >= Config.MinimumSpeed_Mps);
MotionTimer(IN := Comparable, PT := T#1h);
StopTimer(IN := Stopping, PT := T#1h);
IF NOT Comparable THEN StartCapturedM1:=FALSE; StartCapturedM2:=FALSE; ReleaseMsM1:=0; ReleaseMsM2:=0; ApplyMsM1:=0; ApplyMsM2:=0; END_IF;
IF Comparable AND (M1Speed_Mps >= Config.MinimumSpeed_Mps) AND NOT StartCapturedM1 THEN StartMsM1:=TIME_TO_UDINT(MotionTimer.ET); StartCapturedM1:=TRUE; END_IF;
IF Comparable AND (M2Speed_Mps >= Config.MinimumSpeed_Mps) AND NOT StartCapturedM2 THEN StartMsM2:=TIME_TO_UDINT(MotionTimer.ET); StartCapturedM2:=TRUE; END_IF;
{endregion}

{region "§2 Mesure symétrie"}
IF Qualified THEN
    IF M1BrakeCmd AND M1BrakeApplied THEN ReleaseMsM1 := ReleaseMsM1 + REAL_TO_UDINT(CycleTime.CycleTimeS * 1000.0); END_IF;
    IF M2BrakeCmd AND M2BrakeApplied THEN ReleaseMsM2 := ReleaseMsM2 + REAL_TO_UDINT(CycleTime.CycleTimeS * 1000.0); END_IF;
    IF NOT M1BrakeCmd AND NOT M1BrakeApplied THEN ApplyMsM1 := ApplyMsM1 + REAL_TO_UDINT(CycleTime.CycleTimeS * 1000.0); END_IF;
    IF NOT M2BrakeCmd AND NOT M2BrakeApplied THEN ApplyMsM2 := ApplyMsM2 + REAL_TO_UDINT(CycleTime.CycleTimeS * 1000.0); END_IF;
    IF SyncDeviation_M > Data.MaxSyncDeviation_M THEN Data.MaxSyncDeviation_M := SyncDeviation_M; END_IF;
END_IF;
IF PreviousQualified AND NOT Comparable THEN Stopping:=TRUE; StopCapturedM1:=FALSE; StopCapturedM2:=FALSE; StopStartM1_M:=M1Position_M; StopStartM2_M:=M2Position_M; END_IF;
IF Stopping THEN
    IF (M1Speed_Mps < Config.MinimumSpeed_Mps) AND NOT StopCapturedM1 THEN StopMsM1:=TIME_TO_UDINT(StopTimer.ET); StopCapturedM1:=TRUE; END_IF;
    IF (M2Speed_Mps < Config.MinimumSpeed_Mps) AND NOT StopCapturedM2 THEN StopMsM2:=TIME_TO_UDINT(StopTimer.ET); StopCapturedM2:=TRUE; END_IF;
    IF StopCapturedM1 AND StopCapturedM2 THEN
        Data.DeltaStartDelay_Ms := DINT_TO_UDINT(ABS(UDINT_TO_DINT(StartMsM1) - UDINT_TO_DINT(StartMsM2)));
        Data.DeltaBrakeReleaseTime_Ms := DINT_TO_UDINT(ABS(UDINT_TO_DINT(ReleaseMsM1) - UDINT_TO_DINT(ReleaseMsM2)));
        Data.DeltaBrakeApplyTime_Ms := DINT_TO_UDINT(ABS(UDINT_TO_DINT(ApplyMsM1) - UDINT_TO_DINT(ApplyMsM2)));
        Data.DeltaStopDistance_Mm := REAL_TO_UDINT(ABS(ABS(M1Position_M - StopStartM1_M) - ABS(M2Position_M - StopStartM2_M)) * 1000.0);
        Data.DeltaStopTime_Ms := DINT_TO_UDINT(ABS(UDINT_TO_DINT(StopMsM1) - UDINT_TO_DINT(StopMsM2))); Stopping := FALSE; SymmetryValid := TRUE;
    END_IF;
END_IF;
{endregion}

{region "§3 Sortie"}
SymmetryOk := SymmetryValid AND (Data.DeltaStartDelay_Ms<=Config.DeltaStartDelay_Ms) AND (Data.DeltaBrakeReleaseTime_Ms<=Config.DeltaBrakeReleaseTime_Ms) AND (Data.DeltaBrakeApplyTime_Ms<=Config.DeltaBrakeApplyTime_Ms) AND (Data.DeltaStopDistance_Mm<=Config.DeltaStopDistance_Mm) AND (Data.DeltaStopTime_Ms<=Config.DeltaStopTime_Ms);
PreviousQualified := Qualified;
{endregion}

(* ---- FB_WinchCmdArbitrationM1.st ---- *)
(* ═══════════════════════════════════════════════════════════════
   🪝 FB_WinchCmdArbitrationM1 — Arbitrage de commande treuil M1
   ───────────────────────────────────────────────────────────────
   🎯 Rôle : Arbitrer la source de commande M1 (joystick / boutons IHM /
       demande cycle selon le mode) et produire la commande arbitrée.
   🔌 FB d'arbitrage (non-mouvement) : ne porte ni SafeStop ni StartStop
       de sécurité — il produit la commande logique, la safety reste dans
       FB_Safety_Winch / FB_Winch.
   📄 Doc : DOC/AF/AF_Partie-10_Fonction_Winch_v2.1.md
   🔒 Bit-identique à l'ancien PRG_04 §3 (refactor POO).
   🪜 -B : la sortie est désormais un PALIER (StepTgt, 1-5) au lieu d'un
       pourcentage. En SEMI_AUTO, passthrough de ReqWinch.StepTgt ; en manuel,
       le joystick est le producteur UNIQUE du palier (passthrough de
       Joystick.AxisY.StepTgt), boutons/both = palier 5 (pleine vitesse).
   ═══════════════════════════════════════════════════════════════ *)

FUNCTION_BLOCK FB_WinchCmdArbitrationM1
VAR_INPUT
    Enable     : BOOL;  // --> [CMD] Autorisation FB (TRUE=arbitre actif)
    Joystick   : ST_AcquisitionJoystickQualified;  // --> [HW] Données joystick qualifiées (AxisY, DeadmanArmed)
    Auth       : ST_Modes_Autorisations;          // --> [CMD] Autorisations mode (Mode, JoystickWinchSelectArbitrated)
    ReqWinch   : ST_ProgramWinchRequest;            // --> [REQ] Demande cycle treuil M1 (SEMI_AUTO)
    BothIntent : ST_WinchBothIntent;           // --> [CMD] Intention both opérateur (source unique PRG_03)
    IHM        : ST_fbWinchCmdArbitration_IHM;  // --> [CMD] Boutons IHM (BtnAscentM1/BtnDescentM1, both)
    TglJoystickMaster : BOOL;  // --> [CMD] Toggle joystick maître global (Modes.Cmd, source unique)
    Context    : ST_fbWinchCmdArbitration_Context; // --> [STAT] Gating benne/synchro (partagé M1/M2)
    Cfg        : ST_fbWinchCmdArbitration_Cfg;     // --> [CFG] Palier boutons/both (BtnStepTgt)
END_VAR
VAR_OUTPUT
    Ready     : BOOL;  // <-- [STAT] FB prêt à arbitrer (Enable)
    RunRequest : BOOL; // <-- [CMD] Demande marche arbitrée
    ReqAscent  : BOOL; // <-- [CMD] Demande montée arbitrée
    ReqDescend : BOOL; // <-- [CMD] Demande descente arbitrée
    StepTgt   : INT;   // <-- [CMD] Palier de vitesse arbitré (1..5, 0 = arrêt)
END_VAR
VAR
    BenneBusyFallEdge : F_TRIG;  // . [LOC] Front descendant action benne (arrêt forcé)
    BothDirectionAuthorized : BOOL; // . [LOC] Atomicité Both : deux axes autorisés dans le même sens
    RequestConflict         : BOOL; // . [LOC] Double demande de sens refusée
END_VAR

// === IMPLEMENTATION ===

Ready := Enable;

// Front de fin d'action benne (détecté en interne, mécanisme de sécurité)
BenneBusyFallEdge(CLK := Context.BucketBusy);

IF NOT Enable THEN
    RunRequest := FALSE;
    ReqAscent  := FALSE;
    ReqDescend := FALSE;
    StepTgt   := 0;
ELSE
    // ── Pont SEMI_AUTO : consomme la demande du séquenceur de cycle ──
    IF Auth.Mode = E_Mode.SEMI_AUTO THEN
        // Axe X translation prioritaire : aucun contacteur treuil pendant un jog X.
        RunRequest := ReqWinch.RunRequest AND (Joystick.AxisX.Direction = 0);
        ReqAscent  := ReqWinch.ReqAscent;
        ReqDescend := ReqWinch.ReqDescend;
        StepTgt   := ReqWinch.StepTgt;
    ELSE
        // ── Mode manuel : commande both issue de l'intention UNIQUE PRG_03 (BothIntent),
        //    commande unitaire M1 dérivée des boutons/joystick (Select=1). ──
        // 🪜 StepTgt : le joystick est le producteur UNIQUE du palier (FB_Joystick §6).
        //    Boutons/both = pleine vitesse (100 % → palier 5) ; joystick = passthrough
        //    de Joystick.AxisY.StepTgt. Plus de re-dérivation %→palier ici.
        IF NOT TglJoystickMaster THEN
            // Mode Boutons IHM
            IF BothIntent.Active THEN
                // Both (BtnWinchBothAscent/Descent) — source unique PRG_03, plus de re-dérivation
                ReqAscent  := BothIntent.ReqAscent;
                ReqDescend := BothIntent.ReqDescend;
                StepTgt   := Cfg.BtnStepTgt;   // 100 % → palier max (configurable)
            ELSIF IHM.BtnAscentM1 THEN
                ReqAscent  := TRUE;
                ReqDescend := FALSE;
                StepTgt   := Cfg.BtnStepTgt;
            ELSIF IHM.BtnDescentM1 THEN
                ReqAscent  := FALSE;
                ReqDescend := TRUE;
                StepTgt   := Cfg.BtnStepTgt;
            ELSE
                ReqAscent  := FALSE;
                ReqDescend := FALSE;
                StepTgt   := 0;
            END_IF;
        ELSE
            // Mode Joystick Maître — M1 unitaire si Select = 1, both si Select = 0
            IF Auth.JoystickWinchSelectArbitrated = 1 THEN
                ReqAscent  := Joystick.AxisY.Direction > 0;
                ReqDescend := Joystick.AxisY.Direction < 0;
                StepTgt   := Joystick.AxisY.StepTgt;
            ELSIF BothIntent.Active THEN
                // Both (Select=0) — source unique PRG_03, plus de re-dérivation
                ReqAscent  := BothIntent.ReqAscent;
                ReqDescend := BothIntent.ReqDescend;
                StepTgt   := Joystick.AxisY.StepTgt;
            ELSE
                ReqAscent  := FALSE;
                ReqDescend := FALSE;
                StepTgt   := 0;
            END_IF;
        END_IF;

        // Gating StartStop (bit-identique PRG_04 §3) — homme-mort qualifié en joystick
        // 🔗 Atomicité Both : en commande both, la commande ne consomme QUE le
        // permit agrégé (BothAscentPermit/BothDescendPermit) du sens demandé — jamais
        // un permit individuel. Si l'un des 2 treuils n'a pas son permit effectif,
        // AUCUN des deux ne part (départ jamais isolé). En unitaire (BothIntent inactif),
        // le gate est neutre.
        RequestConflict := ReqAscent AND ReqDescend;
        BothDirectionAuthorized := (NOT BothIntent.Active)
            OR ((ReqAscent AND NOT ReqDescend) AND Context.M1AscentAllowed AND Context.M2AscentAllowed)
            OR ((ReqDescend AND NOT ReqAscent) AND Context.M1DescendAllowed AND Context.M2DescendAllowed);
        RunRequest := (ReqAscent OR ReqDescend) AND NOT RequestConflict
                  AND NOT Context.BucketBusy
                  AND NOT Context.WinchBothMotionBlockedByBucket
                  AND NOT ((Context.SyncBlocksAscent   AND ReqAscent)
                        OR (Context.SyncBlocksDescent AND ReqDescend))
                  AND (NOT TglJoystickMaster OR Joystick.DeadmanArmed)
                  // Interlock inter-axes : le jog X translation est prioritaire;
                  // aucun treuil joystick ne part avec X encore deflechi.
                  AND (NOT TglJoystickMaster OR (Joystick.AxisX.Direction = 0))
                  AND BothDirectionAuthorized;
    END_IF;

    // Front de fin d'action benne : arrêt forcé sauf mouvement both actif
    IF BenneBusyFallEdge.Q AND NOT (BothIntent.Active AND (BothIntent.ReqAscent OR BothIntent.ReqDescend)) THEN
        RunRequest := FALSE;
    END_IF;
END_IF;

END_FUNCTION_BLOCK

(* ---- FB_WinchCmdArbitrationM2.st ---- *)
(* ═══════════════════════════════════════════════════════════════
   🪝 FB_WinchCmdArbitrationM2 — Arbitrage de commande treuil M2
   ───────────────────────────────────────────────────────────────
   🎯 Rôle : Arbitrer la source de commande M2 (joystick / boutons IHM /
       demande cycle / chemin benne selon le mode) et produire la commande arbitrée.
   🔌 FB d'arbitrage (non-mouvement) : ne porte ni SafeStop ni StartStop
       de sécurité — il produit la commande logique, la safety reste dans
       FB_Safety_Winch / FB_Winch.
   📄 Doc : DOC/AF/AF_Partie-10_Fonction_Winch_v2.1.md
   🔒 Bit-identique à l'ancien PRG_04 §3 (refactor POO).
   ⚠️ Asymétries M2 vs M1 : chemin benne (override), Select=0/2, synchro inversée.
   🪜 -B : la sortie est désormais un PALIER (StepTgt, 1-5) au lieu d'un
       pourcentage. En SEMI_AUTO, passthrough de ReqWinch.StepTgt ; en manuel,
       le joystick est le producteur UNIQUE du palier (passthrough de
       Joystick.AxisY.StepTgt), boutons/both = palier 5, override benne = palier
       joystick borne par le plafond de configuration.
   ═══════════════════════════════════════════════════════════════ *)

FUNCTION_BLOCK FB_WinchCmdArbitrationM2
VAR_INPUT
    Enable     : BOOL;  // --> [CMD] Autorisation FB (TRUE=arbitre actif)
    Joystick   : ST_AcquisitionJoystickQualified;  // --> [HW] Données joystick qualifiées (AxisY, DeadmanArmed)
    Auth       : ST_Modes_Autorisations;          // --> [CMD] Autorisations mode (Mode, JoystickWinchSelectArbitrated)
    ReqWinch   : ST_ProgramWinchRequest;            // --> [REQ] Demande cycle treuil M2 (SEMI_AUTO)
    BothIntent : ST_WinchBothIntent;           // --> [CMD] Intention both opérateur (source unique PRG_03)
    IHM        : ST_fbWinchCmdArbitration_IHM;  // --> [CMD] Boutons IHM (BtnAscentM2/BtnDescentM2, both)
    TglJoystickMaster : BOOL;  // --> [CMD] Toggle joystick maître global (Modes.Cmd, source unique)
    Context    : ST_fbWinchCmdArbitration_Context; // --> [STAT] Gating benne/synchro + chemin benne (partagé M1/M2)
    Cfg        : ST_fbWinchCmdArbitration_Cfg;     // --> [CFG] Vitesse override benne
END_VAR
VAR_OUTPUT
    Ready     : BOOL;  // <-- [STAT] FB prêt à arbitrer (Enable)
    RunRequest : BOOL; // <-- [CMD] Demande marche arbitrée
    ReqAscent  : BOOL; // <-- [CMD] Demande montée arbitrée
    ReqDescend : BOOL; // <-- [CMD] Demande descente arbitrée
    StepTgt   : INT;   // <-- [CMD] Palier de vitesse arbitré (1..5, 0 = arrêt)
END_VAR
VAR
    BenneBusyFallEdge : F_TRIG;  // . [LOC] Front descendant action benne (arrêt forcé)
    BothDirectionAuthorized : BOOL; // . [LOC] Atomicité Both : deux axes autorisés dans le même sens
    RequestConflict         : BOOL; // . [LOC] Double demande de sens refusée
    BucketRequestedStep     : INT;  // . [LOC] Palier joystick benne avant plafond de configuration
END_VAR

// === IMPLEMENTATION ===

Ready := Enable;

// Front de fin d'action benne (détecté en interne, mécanisme de sécurité)
BenneBusyFallEdge(CLK := Context.BucketBusy);

IF NOT Enable THEN
    RunRequest := FALSE;
    ReqAscent  := FALSE;
    ReqDescend := FALSE;
    StepTgt   := 0;
ELSE
    // ── Chemin benne : M2 piloté par l'action benne (override) ──
    // ⚠️ SÉCURITÉ : l'override benne ne s'applique QUE là où la benne est censée
    // bouger seule (M2 relatif à M1) : jog benne unitaire (WinchSel=2) ou cycle
    // AUTO/SEMI_AUTO qui séquence la benne délibérément. En pilotage COUPLÉ manuel
    // (WinchSel=0) ou unitaire M1 (WinchSel=1), une benne restée Busy NE DOIT PAS
    // détourner M2 : sinon M2 suit la benne pendant que M1 suit le both-intent
    // -> câbles désynchronisés (REX MES 2026-09-04, quasi-casse machine).
    IF Context.BucketBusy AND Context.BucketM2RunRequest
       AND ((Auth.JoystickWinchSelectArbitrated = 2)
            OR (Auth.Mode = E_Mode.SEMI_AUTO)) THEN
        // Axe X translation prioritaire : aucun contacteur treuil pendant un jog X.
        RunRequest := Context.BucketM2RunRequest AND (Joystick.AxisX.Direction = 0);
        ReqAscent  := Context.BucketM2ReqAscent;
        ReqDescend := Context.BucketM2ReqDescend;
        // Le plafond benne borne la consigne joystick ; il ne la remplace pas.
        BucketRequestedStep := LIMIT(1, Joystick.AxisY.StepTgt, 5);
        IF ReqDescend THEN
            StepTgt := MIN(BucketRequestedStep, Cfg.BucketOverrideStepDownTgt);
        ELSIF ReqAscent AND Context.BucketHandoffP1Active THEN
            StepTgt := 1;
        ELSIF ReqAscent AND Context.BucketAutoCloseActive THEN
            StepTgt := MIN(BucketRequestedStep, Cfg.BucketAutoMaxStepUp);
        ELSE
            StepTgt := MIN(BucketRequestedStep, Cfg.BucketOverrideStepUpTgt);
        END_IF;
    ELSE
        // ── Pont SEMI_AUTO : consomme la demande du séquenceur de cycle ──
        IF Auth.Mode = E_Mode.SEMI_AUTO THEN
            // Axe X translation prioritaire : aucun contacteur treuil pendant un jog X.
            RunRequest := ReqWinch.RunRequest AND (Joystick.AxisX.Direction = 0);
            ReqAscent  := ReqWinch.ReqAscent;
            ReqDescend := ReqWinch.ReqDescend;
            StepTgt   := ReqWinch.StepTgt;
        ELSE
            // ── Mode manuel : commande both issue de l'intention UNIQUE PRG_03 (BothIntent),
            //    commande unitaire M2 dérivée des boutons/joystick (Select=2). ──
            // 🪜 StepTgt : le joystick est le producteur UNIQUE du palier (FB_Joystick §6).
            //    Boutons/both = pleine vitesse (100 % → palier 5) ; joystick = passthrough
            //    de Joystick.AxisY.StepTgt. Plus de re-dérivation %→palier ici.
            IF NOT TglJoystickMaster THEN
                // Mode Boutons IHM
                IF BothIntent.Active THEN
                    // Both (BtnWinchBothAscent/Descent) — source unique PRG_03, plus de re-dérivation
                    ReqAscent  := BothIntent.ReqAscent;
                    ReqDescend := BothIntent.ReqDescend;
                    StepTgt   := Cfg.BtnStepTgt;   // 100 % → palier max (configurable)
                ELSIF IHM.BtnAscentM2 THEN
                    ReqAscent  := TRUE;
                    ReqDescend := FALSE;
                    StepTgt   := Cfg.BtnStepTgt;
                ELSIF IHM.BtnDescentM2 THEN
                    ReqAscent  := FALSE;
                    ReqDescend := TRUE;
                    StepTgt   := Cfg.BtnStepTgt;
                ELSE
                    ReqAscent  := FALSE;
                    ReqDescend := FALSE;
                    StepTgt   := 0;
                END_IF;
            ELSE
                // Mode Joystick Maître — M2 unitaire si Select = 2, both si Select = 0
                IF Auth.JoystickWinchSelectArbitrated = 2 THEN
                    ReqAscent  := Joystick.AxisY.Direction > 0;
                    ReqDescend := Joystick.AxisY.Direction < 0;
                    StepTgt   := Joystick.AxisY.StepTgt;
                ELSIF BothIntent.Active THEN
                    // Both (Select=0) — source unique PRG_03, plus de re-dérivation
                    ReqAscent  := BothIntent.ReqAscent;
                    ReqDescend := BothIntent.ReqDescend;
                    StepTgt   := Joystick.AxisY.StepTgt;
                ELSE
                    ReqAscent  := FALSE;
                    ReqDescend := FALSE;
                    StepTgt   := 0;
                END_IF;
            END_IF;

            // Gating StartStop (bit-identique PRG_04 §3) — synchro INVERSÉE vs M1,
            // homme-mort qualifié en joystick
            // 🔗 Atomicité Both : cf. M1 — en both, la commande ne consomme QUE le
            // permit agrégé du sens demandé. Départ jamais isolé entre les 2 treuils.
            RequestConflict := ReqAscent AND ReqDescend;
            BothDirectionAuthorized := (NOT BothIntent.Active)
                OR ((ReqAscent AND NOT ReqDescend) AND Context.M1AscentAllowed AND Context.M2AscentAllowed)
                OR ((ReqDescend AND NOT ReqAscent) AND Context.M1DescendAllowed AND Context.M2DescendAllowed);
            RunRequest := (ReqAscent OR ReqDescend) AND NOT RequestConflict
                      AND NOT Context.WinchBothMotionBlockedByBucket
                      AND NOT ((Context.SyncBlocksAscent   AND ReqDescend)
                            OR (Context.SyncBlocksDescent AND ReqAscent))
                      AND (NOT TglJoystickMaster OR Joystick.DeadmanArmed)
                      // Interlock inter-axes : le jog X translation est prioritaire;
                      // aucun treuil joystick ne part avec X encore deflechi.
                      AND (NOT TglJoystickMaster OR (Joystick.AxisX.Direction = 0))
                      AND BothDirectionAuthorized;
        END_IF;
    END_IF;

    // Front de fin d'action benne : arrêt forcé sauf mouvement both actif
    IF BenneBusyFallEdge.Q AND NOT (BothIntent.Active AND (BothIntent.ReqAscent OR BothIntent.ReqDescend)) THEN
        RunRequest := FALSE;
    END_IF;
END_IF;

END_FUNCTION_BLOCK

(* ---- FB_WinchDirectionInterlock.st ---- *)
(* =======================================================================
   🔀 FB_WinchDirectionInterlock — Interlock de changement de sens
   ───────────────────────────────────────────────────────────────
   🎯 Rôle : Temporise l'INVERSION de sens d'un treuil, en creditant le
             temps d'arret physique reel deja ecoule (dead time)
   📄 Doc métier : DOC/AF/AF_Partie-10_Fonction_Winch_v2.1.md
   🔌 Interface : Brique technique (contrat light, pas de defaut)
   🔒 Sécurité : D18 — au front montant Enable, n'adopte pas le sens
                 immediatement (temps mort) ; pas de redemarrage inrush.
                 Le sens IDENTIQUE au dernier sens adopte reste toujours
                 immediat depuis le neutre : seule l'INVERSION est temporisee.
                 Purge de DeadTimeArmed garantie des que le temps mort est
                 ecoule (T325 phase 1). Limite residuelle connue (T325
                 phase 2, non couverte ici) : si la demande redevient le
                 MEME sens que le dernier commande alors que DeadTimeArmed
                 vient d'etre arme, DirectionChanged reste FALSE et le
                 temps mort ne peut jamais etre mesure -- seule sortie
                 encore possible dans ce cas precis : retour au neutre ou
                 Reset.
   ======================================================================= *)

FUNCTION_BLOCK PUBLIC FB_WinchDirectionInterlock
VAR_INPUT
    Enable          : BOOL;   // --> [CMD] Gate TON (TRUE = treuil arrete, contacteurs retombes)
    EnableRising    : BOOL;   // --> [CMD] Front montant Enable du FB parent (D18)
    Reset           : BOOL;   // --> [CMD] Acquittement defaut (front) : purge la memoire de direction
    ReqAscent       : BOOL;   // --> [CMD] Demande montée
    ReqDescend      : BOOL;   // --> [CMD] Demande descente
    ChangeDelayAscent   : TIME;   // --> [CFG] Delai interlock changement de sens montee
    ChangeDelayDescent : TIME;   // --> [CFG] Delai interlock changement de sens descente
END_VAR
VAR_OUTPUT
    CommandedAscent         : BOOL;  // <-- [DIAG] Sens interne mémorisé : montée
    CommandedDescend        : BOOL;  // <-- [DIAG] Sens interne mémorisé : descente
    RequestConflict         : BOOL;  // <-- [DIAG] Double demande refusée
    DirectionChangePending  : BOOL;  // <-- [DIAG] Changement de sens en attente
    DelayElapsed            : TIME;  // <-- [DIAG] Ecoule delai changement de sens
END_VAR
VAR
    DirectionChangeDelay  : TON;      // . [LOC] Xa->Xb : compte le reliquat apres la nouvelle demande d'inversion
    StoppedTimer          : TON;      // . [LOC] Xc->Xd : accumule le temps d'arret physique reel (Enable, hors demande)
    CapturedStoppedTime   : TIME;     // . [LOC] Arret reel credite, fige au front RequestActive, purge une fois consomme
    RemainingDelay        : TIME;     // . [LOC] Reliquat a appliquer par DirectionChangeDelay (delai plein - arret credite)
    EffectiveDelay        : TIME;     // . [LOC] Delai plein selon sens demande
    MaxDirectionDelay     : TIME;     // . [LOC] MAX(ChangeDelayAscent, ChangeDelayDescent) : base d'accumulation StoppedTimer
    DeadTimeArmed         : BOOL;     // . [LOC] Temps mort D18 arme (front Enable)
    LastAscent            : BOOL;     // . [LOC] Dernier sens adopté : montée
    LastDescend           : BOOL;     // . [LOC] Dernier sens adopté : descente
    RequestActive         : BOOL;     // . [LOC] Une seule demande de sens active
    RequestActiveRising   : R_TRIG;   // . [LOC] Front nouvelle demande : capture le credit avant le rappel de StoppedTimer
    DirectionChanged      : BOOL;     // . [LOC] Demande différente du sens commandé
    ResetEdge             : R_TRIG;   // . [LOC] Front Reset : purge la memoire de direction
END_VAR

// === IMPLEMENTATION ===

// Front Reset : purge la memoire de direction (un acquittement conscient reinitialise
// l'historique, une reprise apres Reset est un depart propre, pas une inversion).
ResetEdge(CLK := Reset);
IF ResetEdge.Q THEN
    LastAscent := FALSE;
    LastDescend := FALSE;
    CommandedAscent := FALSE;
    CommandedDescend := FALSE;
    DeadTimeArmed := FALSE;
    DirectionChangePending := FALSE;
    CapturedStoppedTime := T#0ms;
END_IF;

RequestConflict := ReqAscent AND ReqDescend;
RequestActive := (ReqAscent OR ReqDescend) AND NOT RequestConflict;

// Xc->Xd : capture l'arret physique REEL deja ecoule (StoppedTimer.ET) AU FRONT de
// la nouvelle demande, AVANT le rappel de StoppedTimer plus bas dans ce scan (un TON
// dont IN retombe a FALSE remet son ET a 0 des cet appel — lire apres serait deja 0).
RequestActiveRising(CLK := RequestActive);
IF RequestActiveRising.Q THEN
    CapturedStoppedTime := StoppedTimer.ET;
END_IF;

// Délai plein selon le sens demandé, et base commune pour l'accumulation d'arret
// (le sens final n'est pas encore connu pendant le neutre).
IF ReqAscent AND NOT ReqDescend THEN
    EffectiveDelay := ChangeDelayAscent;
ELSE
    EffectiveDelay := ChangeDelayDescent;
END_IF;
MaxDirectionDelay := MAX(ChangeDelayAscent, ChangeDelayDescent);
// Comparaison AVANT soustraction : TIME est un DWORD non signe cote CODESYS, une
// soustraction dont le resultat mathematique serait negatif (ex: T#500ms - T#800ms)
// deborde silencieusement vers ~T#49j au lieu de saturer a 0 -- MAX(..., T#0ms)
// APRES une soustraction debordee ne corrige rien (le DWORD deborde reste "positif").
IF CapturedStoppedTime >= EffectiveDelay THEN
    RemainingDelay := T#0ms;
ELSE
    RemainingDelay := EffectiveDelay - CapturedStoppedTime;
END_IF;

DirectionChanged := (ReqAscent AND NOT CommandedAscent)
                 OR (ReqDescend AND NOT CommandedDescend)
                 OR (CommandedAscent AND NOT ReqAscent)
                 OR (CommandedDescend AND NOT ReqDescend);

// D18 : au front montant Enable avec sens maintenu, armer le temps mort
// (ne pas re-adopter le sens immediatement — pas de redemarrage inrush).
IF EnableRising AND RequestActive THEN
    DeadTimeArmed := TRUE;
END_IF;

// Xc->Xd : StoppedTimer compte l'arret physique REEL (Enable = treuil arrete,
// contacteurs retombes, cf. FB_Winch) pendant TOUT le neutre, jamais reinitialise
// par le simple relachement du joystick — c'est ce cumul qui alimente la capture
// ci-dessus au scan suivant.
StoppedTimer(IN := Enable AND NOT RequestActive, PT := MaxDirectionDelay);

// Xa->Xb : compte le reliquat (delai plein - arret deja credite) apres la nouvelle
// demande d'inversion.
DirectionChangeDelay(
    IN := Enable AND RequestActive AND DirectionChanged,
    PT := RemainingDelay
);
DelayElapsed := DirectionChangeDelay.ET;

// Adoption du sens
IF NOT RequestActive THEN
    // Neutre ou double demande : aucun sens commandé. Une double demande est
    // explicitement refusée, sans priorité implicite.
    CommandedAscent := FALSE;
    CommandedDescend := FALSE;
    DirectionChangePending := FALSE;
    DeadTimeArmed := FALSE;
ELSIF DirectionChangeDelay.Q THEN
    // Temps mort ecoule : adoption du sens, y compris si DeadTimeArmed etait pose
    // (purge desormais atteignable -- le temps mort minimal a ete respecte, il ne
    // doit pas rester arme indefiniment une fois le delai reellement ecoule).
    CommandedAscent := ReqAscent;
    CommandedDescend := ReqDescend;
    DirectionChangePending := FALSE;
    DeadTimeArmed := FALSE;
ELSIF DeadTimeArmed THEN
    // D18 : temps mort au front Enable — pas d'adoption immediate tant que le
    // delai (ci-dessus) n'est pas ecoule.
    DirectionChangePending := TRUE;
ELSIF NOT (CommandedAscent OR CommandedDescend) THEN
    // Depuis le neutre : depart immediat si reprise du MEME sens (ou premier sens),
    // sinon (sens oppose) pending + delai dedie obligatoire.
    IF (NOT (LastAscent OR LastDescend))
       OR (ReqAscent AND LastAscent)
       OR (ReqDescend AND LastDescend) THEN
        CommandedAscent := ReqAscent;
        CommandedDescend := ReqDescend;
        DirectionChangePending := FALSE;
    ELSE
        DirectionChangePending := TRUE;
    END_IF;
ELSIF DirectionChanged THEN
    // Inversion directe (sans passage au neutre) : pending + delai
    DirectionChangePending := TRUE;
ELSE
    DirectionChangePending := FALSE;
END_IF;

// Memorise le dernier sens non nul ADOPTE (pas la simple demande) : c'est ce sens qui
// sert de reference pour detecter une reprise opposee apres passage au neutre.
IF CommandedAscent OR CommandedDescend THEN
    LastAscent := CommandedAscent;
    LastDescend := CommandedDescend;
END_IF;

// Le sens adopte correspond desormais a la demande (aucune inversion en cours) :
// le credit d'arret est CONSOMME. Une inversion ULTERIEURE sans nouveau passage au
// neutre (RequestActive reste continuellement vrai) ne doit jamais reutiliser un
// arret perime — elle applique alors le delai plein (CapturedStoppedTime := 0).
IF NOT DirectionChangePending AND (CommandedAscent = ReqAscent) AND (CommandedDescend = ReqDescend) THEN
    CapturedStoppedTime := T#0ms;
END_IF;

END_FUNCTION_BLOCK

(* ---- FB_WinchLoadEstimator.st ---- *)
(* =======================================================================
   📊 FB_WinchLoadEstimator — Estimation empirique de charge treuil
   ───────────────────────────────────────────────────────────────
   🎯 Rôle : Estimation informative de la charge par croisement palier/vitesse
   📄 Doc métier : DOC/AF/AF_Partie-10_Fonction_Winch_v2.1.md
   🔌 Interface : Brique de diagnostic/mesure (1 instance par treuil)
   🔒 Sécurité : Aucune commande moteur ni action sur SafeStop (information IHM)
   ======================================================================= *)

FUNCTION_BLOCK PUBLIC FB_WinchLoadEstimator

VAR_INPUT
    // === COMMANDES ET CONSIGNES ===
    Enable                          : BOOL;                           // --> [CMD] Autorisation generale FB
    Reset                           : BOOL;                           // --> [CMD] Acquittement defaut sur front
    Mode                            : E_Mode;                         // --> [CMD] Mode d'exploitation actif
    ActiveSpeedStep                 : INT;                            // --> [CMD] Palier commande actif (0..5)

    // === SECOURS ET HARDWARE ===
    PowerContactorEngaged           : BOOL;                           // --> [SAFE] Chaine AU rearmee et puissance OK
    MeasuredSpeedMps                : REAL;                           // --> [HW] Vitesse cable absolue (m/s)
    MeasuredSpeedSignedMps          : REAL;                           // --> [HW] Vitesse signee (+: montee, -: descente) (m/s)

    // === REGLAGES ET TABLES ===
    SpeedConfig                     : ST_fbWinchLoadEstimator_SpeedCfg;            // --> [CFG] Configuration des plages de vitesse
    LoadTable                       : ST_fbWinchLoadEstimator_Table;      // --> [CFG] Table empirique d'estimation 5x5
END_VAR
VAR_OUTPUT
    // === ETATS IEC ET SYNOPTIQUE ===
    Ready                           : BOOL;                           // <-- [STAT] FB pret a fonctionner
    // 🧩 Statut transverse (forme cible ST_Fault)
    Fault                           : ST_Fault;

    // === DIAGNOSTICS ET ESTIMATIONS ===
    SpeedBand                       : INT;                            // <-- [DIAG] Bande de vitesse courante (0..5)
    EstimatedLoadPct                : REAL;                           // <-- [DIAG] Estimation de charge (0..100%)
    Configured                      : BOOL;                           // <-- [STAT] Table explicitement validee
    Ascending                       : BOOL;                           // <-- [STAT] Ascending effective mesuree en cours
END_VAR
VAR
    // === DETECTEURS ET TIMERS INTERNES ===
    ResetEdge                       : R_TRIG;                         // . [LOC] Detecteur front montant Reset

    // === VARIABLES LOCALES CALCULÉES ===
    PreviousSpeedBand               : INT;                            // . [LOC] Memoire bande de vitesse cycle precedent
    HasPreviousBand                 : BOOL;                           // . [LOC] Indicateur premiere bande memorisee
    SelectedLoadPct                 : REAL;                           // . [LOC] Valeur de charge extraite de la table
    ConfigOrSpeedFault              : BOOL;                           // . [LOC] Latch défaut configuration / vitesse

    // === SOCLE DEFAUT ===
    instFault                       : FB_FaultCore;                   // * [INST] Socle défaut transverse
    instCauses                      : ARRAY[0..15] OF ST_FaultCause;  // . [LOC] Table des causes nommées
END_VAR

// === IMPLEMENTATION ===

{region "§1 Causes & Socle Défaut (évalué en continu)"}
// 🔑 1. FRONTS
ResetEdge(CLK := Reset);

IF ResetEdge.Q AND (MeasuredSpeedMps >= 0.0) THEN
    ConfigOrSpeedFault := FALSE;
END_IF;

instCauses[0].Active   := ConfigOrSpeedFault;
instCauses[0].Latching := TRUE;
instCauses[0].Texte    := 'Parametrage ou vitesse estimation charge invalide';

// Appel du socle de défaut
instFault(Enable := Enable, Reset := Reset, Causes := instCauses);
Fault := instFault.Fault;
{endregion}

{region "§2 Gate neutralisation"}
// 🛑 2. GATE
IF NOT Enable OR NOT PowerContactorEngaged THEN
    Ready := FALSE;
    SpeedBand := 0;
    EstimatedLoadPct := 0.0;
    Configured := FALSE;
    Ascending := FALSE;
    HasPreviousBand := FALSE;
    RETURN;
END_IF;

Ready := Enable AND NOT Fault.Latched;
Configured := LoadTable.IsConfigured;
Ascending := (MeasuredSpeedSignedMps > 0.0);
{endregion}

{region "§3 Classement vitesse"}
// 📏 3. CLASSEMENT DE LA VITESSE — hystérésis autour des 4 frontières.
IF (MeasuredSpeedMps < 0.0) OR (SpeedConfig.MaxMeasuredSpeedMps <= 0.0) THEN
    ConfigOrSpeedFault := TRUE;
    SpeedBand := 0;
ELSIF NOT HasPreviousBand THEN
    IF MeasuredSpeedMps <= SpeedConfig.SpeedBandMaxMps[1] THEN
        PreviousSpeedBand := 1;
    ELSIF MeasuredSpeedMps <= SpeedConfig.SpeedBandMaxMps[2] THEN
        PreviousSpeedBand := 2;
    ELSIF MeasuredSpeedMps <= SpeedConfig.SpeedBandMaxMps[3] THEN
        PreviousSpeedBand := 3;
    ELSIF MeasuredSpeedMps <= SpeedConfig.SpeedBandMaxMps[4] THEN
        PreviousSpeedBand := 4;
    ELSE
        PreviousSpeedBand := 5;
    END_IF;
    HasPreviousBand := TRUE;
    SpeedBand := PreviousSpeedBand;
ELSE
    IF PreviousSpeedBand < 1 OR PreviousSpeedBand > 5 THEN
        PreviousSpeedBand := 1;
        ConfigOrSpeedFault := TRUE;
    END_IF;

    IF PreviousSpeedBand < 5 THEN
        IF MeasuredSpeedMps > (SpeedConfig.SpeedBandMaxMps[PreviousSpeedBand]
                               + SpeedConfig.SpeedBandHysteresisMps) THEN
            PreviousSpeedBand := PreviousSpeedBand + 1;
        END_IF;
    END_IF;
    IF PreviousSpeedBand > 1 THEN
        IF MeasuredSpeedMps < (SpeedConfig.SpeedBandMaxMps[PreviousSpeedBand - 1]
                               - SpeedConfig.SpeedBandHysteresisMps) THEN
            PreviousSpeedBand := PreviousSpeedBand - 1;
        END_IF;
    END_IF;
    SpeedBand := PreviousSpeedBand;
END_IF;
{endregion}

{region "§4 Lecture table"}
// 📊 4. LECTURE TABLE
EstimatedLoadPct := 0.0;
IF Configured THEN
    IF Ascending THEN
        IF ActiveSpeedStep >= 1 THEN
            IF ActiveSpeedStep <= 5 THEN
                IF SpeedBand >= 1 THEN
                    IF SpeedBand <= 5 THEN
                        SelectedLoadPct := LoadTable.LoadPctByStepAndSpeedBand[ActiveSpeedStep][SpeedBand];
                        IF (SelectedLoadPct < 0.0) OR (SelectedLoadPct > 100.0) THEN
                            ConfigOrSpeedFault := TRUE;
                        ELSE
                            EstimatedLoadPct := SelectedLoadPct;
                        END_IF;
                    END_IF;
                END_IF;
            END_IF;
        END_IF;
    END_IF;
END_IF;
{endregion}

END_FUNCTION_BLOCK

(* ---- FB_WinchSpeedLearning.st ---- *)
(* =======================================================================
   💾 FB_WinchSpeedLearning — Collecteur passif vitesse par palier
   ───────────────────────────────────────────────────────────────
   🎯 Rôle : Apprentissage passif des vitesses reelles par palier (RETAIN)
   📄 Doc metier : DOC/AF/AF_Partie-10_Fonction_Winch_v2.1.md
   🔒 Collecteur pur : aucune commande moteur, aucune surveillance survitesse
   ======================================================================= *)

FUNCTION_BLOCK FB_WinchSpeedLearning
VAR_INPUT
    // === CONTRAT LIGHT (Enable) ===
    Enable                          : BOOL;   // --> [CMD] Autorisation generale FB (TRUE=Autorise)
    LearnStart                      : BOOL;   // --> [CMD] Bit IHM lancer apprentissage
    WinchId                         : INT;    // --> [CMD] Axe cible (1=M1, 2=M2)
    ReqAscent                       : BOOL;   // --> [HW] Mesure active montée
    ReqDescend                      : BOOL;   // --> [HW] Mesure active descente
    StepNumber                      : INT;    // --> [HW] Palier actif (1..5)
    MeasuredSpeedMps                : REAL;   // --> [HW] Vitesse mesuree (m/s)
    MeasuredSpeedValid              : BOOL;   // --> [HW] Mesure exploitable
    LoadPresent                     : BOOL;   // --> [HW] Charge presente (TRUE=charge, FALSE=vide)
    StableForLearn                  : BOOL;   // --> [HW] Conditions stables pour apprentissage

    // === REGLAGES & CONFIGURATION ===
    Config                          : ST_fbWinchSpeedLearning_Cfg; // --> [CFG] Enveloppes de plausibilite par palier
END_VAR
VAR_OUTPUT
    // === CONTRAT LIGHT (Ready) ===
    Ready                           : BOOL;   // <-- [STAT] FB pret (Enable)

    // === ETATS & DIAGNOSTIC ===
    Learning                        : BOOL;   // <-- [STAT] Collecte en cours
    TableComplete                   : BOOL;   // <-- [STAT] Table charge ET vide complete
    LampLearn                       : BOOL;   // <-- [STAT] Voyant IHM apprentissage
    CellsFilled                     : INT;    // <-- [DIAG] Nombre de cellules validees
    CellsTotal                      : INT;    // <-- [DIAG] Nombre total de cellules
END_VAR
VAR_IN_OUT
    // === STRUCTURES DE DONNEES PARTAGEES ===
    Table                           : ST_fbWinchSpeedLearning_Table; // <-> [BUS] Table RETAIN apprentissage
END_VAR
VAR
    // === VARIABLES LOCALES CALCULEES ===
    LearnRequested                  : BOOL;   // . [LOC] Bit IHM + Enable
    MeasureUsable                   : BOOL;   // . [LOC] Mesure valide + conditions stables
    SensActive                      : BOOL;   // . [LOC] Un seul sens actif
    SensConflict                    : BOOL;   // . [LOC] Deux sens actifs : collecte interdite
    StepInRange                     : BOOL;   // . [LOC] Palier dans 1..5
    AxeInRange                      : BOOL;   // . [LOC] Axe dans 1..2
    ContextValid                    : BOOL;   // . [LOC] Sens, palier et axe dans le domaine
    CollectAllowed                  : BOOL;   // . [LOC] Conditions de collecte reunies
    SpeedPlausible                  : BOOL;   // . [LOC] Vitesse dans l'enveloppe du palier
    SensIdx                         : INT;    // . [LOC] Index sens (1=montee, 2=descente)
    ChargeIdx                       : INT;    // . [LOC] Index charge (1=vide, 2=charge)
    CurrentCell                     : ST_fbWinchSpeedLearning_Cell; // . [LOC] Cellule courante
    AxeIdx                          : INT;    // . [LOC] Index axe boucle
    SensLoopIdx                     : INT;    // . [LOC] Index sens boucle
    ChargeLoopIdx                   : INT;    // . [LOC] Index charge boucle
    PalierIdx                       : INT;    // . [LOC] Index palier boucle
END_VAR
VAR CONSTANT
    CST_AxeCount                    : INT := 2;   // Nombre d'axes (M1, M2)
    CST_SensCount                   : INT := 2;   // Nombre de sens (ascending, descending)
    CST_ChargeCount                 : INT := 2;   // Nombre d'etats de charge (vide, charge)
    CST_PalierCount                 : INT := 5;   // Nombre de paliers (1..5)
    CST_IdxAscent                : INT := 1;   // Index sens ascending
    CST_IdxDescent               : INT := 2;   // Index sens descending
    CST_IdxVide                     : INT := 1;   // Index charge vide
    CST_IdxCharge                   : INT := 2;   // Index charge presente
END_VAR

{region "§1 Gate et conditions de collecte"}
Ready := Enable;
Learning := FALSE;
LampLearn := FALSE;

// Conditions de collecte scindees (lisibilite Watch, <=3 termes par predicat)
LearnRequested := Enable AND LearnStart;
MeasureUsable := MeasuredSpeedValid AND StableForLearn;
SensConflict := ReqAscent AND ReqDescend;
SensActive := (ReqAscent OR ReqDescend) AND NOT SensConflict;
StepInRange := (StepNumber >= 1) AND (StepNumber <= CST_PalierCount);
AxeInRange := (WinchId >= 1) AND (WinchId <= CST_AxeCount);
ContextValid := SensActive AND StepInRange AND AxeInRange;
CollectAllowed := LearnRequested AND MeasureUsable AND ContextValid;
{endregion}

{region "§2 Collecte passive"}
IF CollectAllowed THEN
    // Index sens et charge
    IF ReqAscent THEN SensIdx := CST_IdxAscent; ELSE SensIdx := CST_IdxDescent; END_IF;
    IF LoadPresent THEN ChargeIdx := CST_IdxCharge; ELSE ChargeIdx := CST_IdxVide; END_IF;

    // Plausibilite : vitesse dans l'enveloppe du palier (borne min/max)
    SpeedPlausible := (MeasuredSpeedMps >= Config.MinSpeedMps[StepNumber])
                      AND (MeasuredSpeedMps <= Config.MaxSpeedMps[StepNumber]);

    CurrentCell := Table.Cell[WinchId, SensIdx, ChargeIdx, StepNumber];
    IF SpeedPlausible THEN
        // Accumulation (moyenne glissante)
        IF CurrentCell.SampleCount = 0 THEN
            CurrentCell.SpeedMps := MeasuredSpeedMps;
            CurrentCell.SampleCount := 1;
        ELSE
            CurrentCell.SpeedMps := (CurrentCell.SpeedMps * UDINT_TO_REAL(CurrentCell.SampleCount) + MeasuredSpeedMps)
                                    / UDINT_TO_REAL(CurrentCell.SampleCount + 1);
            CurrentCell.SampleCount := CurrentCell.SampleCount + 1;
        END_IF;
        CurrentCell.Valid := (CurrentCell.SampleCount >= Config.MinSamples);
    ELSE
        // Valeur hors enveloppe -> cellule invalidee
        CurrentCell.Valid := FALSE;
        CurrentCell.SampleCount := 0;
        CurrentCell.SpeedMps := 0.0;
    END_IF;
    Table.Cell[WinchId, SensIdx, ChargeIdx, StepNumber] := CurrentCell;

    Learning := TRUE;
    LampLearn := TRUE;
END_IF;
{endregion}

{region "§3 Comptage et completude"}
CellsTotal := CST_AxeCount * CST_SensCount * CST_ChargeCount * CST_PalierCount;
CellsFilled := 0;
FOR AxeIdx := 1 TO CST_AxeCount DO
    FOR SensLoopIdx := 1 TO CST_SensCount DO
        FOR ChargeLoopIdx := 1 TO CST_ChargeCount DO
            FOR PalierIdx := 1 TO CST_PalierCount DO
                IF Table.Cell[AxeIdx, SensLoopIdx, ChargeLoopIdx, PalierIdx].Valid THEN
                    CellsFilled := CellsFilled + 1;
                END_IF;
            END_FOR;
        END_FOR;
    END_FOR;
END_FOR;
TableComplete := (CellsFilled >= CellsTotal);
{endregion}
